// FB_HydraulicsControl with a plant: the pump feedback follows the pump enable output one scan later and the oil pressure
// follows the pump (a starter and a pump that work), the suction feedback follows the suction enable. The sensors are healthy.
// bAuto calls OpenBrake() in every scan (the automatic request of MONETcommon), bManual calls ManualBrake(bSwitch) and
// feeds the switch to bBrakeClearing as MAIN of MONETS/MONETN does. tPumpResetPulse is T#0S: the pump starts at once.
// StepStart()/StepTime() measure real time from the start of a step (the block timers run on the system time).
FUNCTION_BLOCK FB_HydraulicsRig
VAR_INPUT
	stIn		: HalfBROT.ST_HydraulicsIn := (bOilLow := TRUE, bOilHigh := TRUE, bOilCold := TRUE, bOilFilterDirty := TRUE, nOilLevel := 8000);
	bClearing	: BOOL;
	bAzLimit	: BOOL;
	bAuto		: BOOL;
	bManual		: BOOL;
	bSwitch		: BOOL;
	bPumpFollows	: BOOL := TRUE;
	bPressure		: BOOL := TRUE;
	bSuctionFollows	: BOOL := TRUE;
	tHydraulicsWatchdog	: TIME := T#140S;
	tSuctionWatchdog	: TIME := T#15S;
	tPressureWatchdog	: TIME := T#30S;
END_VAR
VAR
	fbComm		: FB_NullComm;
	fb			: HalfBROT.FB_HydraulicsControl(comm := fbComm);
	stOut		: HalfBROT.ST_HydraulicsOut;
	tonStep		: TON;
	nScans		: UDINT;
	nStepScans	: UDINT;
END_VAR

METHOD Scan
nScans := nScans + 1;
nStepScans := nStepScans + 1;
IF bPumpFollows THEN
	stIn.bPumpRunning := stOut.bOilPumpEnable;
END_IF
stIn.bOilPressureOK := stIn.bPumpRunning AND bPressure;
IF bSuctionFollows THEN
	stIn.bSuctionRunning := stOut.bOilSuctionEnable;
END_IF
IF bAuto THEN
	fb.OpenBrake();
END_IF
IF bManual THEN
	bClearing := bSwitch;
	fb.ManualBrake(bSwitch := bSwitch);
END_IF
fb(stIn := stIn, bBrakeClearing := bClearing, bAzimuthLimitSwitch := bAzLimit, tHydraulicsWatchdog := tHydraulicsWatchdog,
	tSuctionWatchdog := tSuctionWatchdog, tPressureWatchdog := tPressureWatchdog, tPumpResetPulse := T#0S, stOut := stOut);
tonStep(IN := TRUE, PT := T#1H);
END_METHOD

METHOD StepStart
tonStep(IN := FALSE, PT := T#1H);
nStepScans := 0;
END_METHOD

METHOD StepTime : BOOL
VAR_INPUT
	tTime	: TIME;
END_VAR
StepTime := tonStep.ET >= tTime;
END_METHOD

METHOD SetEnable
VAR_INPUT
	bOn	: BOOL;
END_VAR
fb.Enable := bOn;
END_METHOD

METHOD SetSuction
VAR_INPUT
	bOn	: BOOL;
END_VAR
fb.ManualStartSuction := bOn;
END_METHOD

METHOD SetStopPump
VAR_INPUT
	bOn	: BOOL;
END_VAR
fb.ManualStopPump := bOn;
END_METHOD

END_FUNCTION_BLOCK

(* stored: Version 1.1.0.1, ProductVersion 3.1.4024.15
   POU FB_HydraulicsRig: Id {9e5eff1a-a9b5-53ef-be33-154116ea001f}, SpecialFunc None
   Method Scan: Id {f5cdac0c-d4f0-5b46-bdb5-96ac2875fe99}
   Method StepStart: Id {5b412144-d45d-5751-a8ad-8345070fe72b}
   Method StepTime: Id {f03c8e75-35a6-5eb0-ba58-4b005a03ced1}
   Method SetEnable: Id {3ecaf0ab-3e22-5f48-acee-a7d3bf29c399}
   Method SetSuction: Id {790ae574-875e-5d0d-9039-d261f13890d4}
   Method SetStopPump: Id {b828b65d-e35a-50cf-9c05-942c73d6f13c} *)
